(* IEC 61131-3 sources: llm-plc-st-eval/data/definitivo/gemini-3.1-pro-preview/I4/zero_shot, 3 files *)

(* ---- ejec_1.st ---- *)
```iecst
FUNCTION_BLOCK FB_EstrellaTriangulo
VAR_INPUT
    btnMarcha : BOOL; // Botón de arranque
    btnParo   : BOOL; // Botón de parada (prioridad a la parada)
END_VAR

VAR_OUTPUT
    kM : BOOL; // Contactor principal
    kY : BOOL; // Contactor de estrella
    kD : BOOL; // Contactor de triángulo
END_VAR

VAR
    tonEstrella   : TON; // Temporizador para la fase de estrella (8s)
    tonTransicion : TON; // Temporizador para el tiempo muerto (100ms)
END_VAR

// 1. Lógica del contactor principal (kM)
// Enclavamiento con btnMarcha, se rompe al pulsar btnParo
kM := (btnMarcha OR kM) AND NOT btnParo;

// 2. Temporizadores
// El temporizador de estrella inicia al arrancar el motor (kM = TRUE)
tonEstrella(IN := kM, PT := T#8S);

// El temporizador de transición inicia cuando termina la fase de estrella
tonTransicion(IN := tonEstrella.Q, PT := T#100MS);

// 3. Lógica de los contactores de fase (con enclavamiento mutuo de seguridad)
// kY se activa con kM, se apaga al terminar tonEstrella, y nunca si kD está activo
kY := kM AND NOT tonEstrella.Q AND NOT kD;

// kD se activa al terminar el tiempo muerto, y nunca si kY está activo
kD := kM AND tonTransicion.Q AND NOT kY;

END_FUNCTION_BLOCK
```

(* ---- ejec_2.st ---- *)
```iecst
FUNCTION_BLOCK FB_EstrellaTriangulo
VAR_INPUT
    btnMarcha : BOOL; (* Botón de inicio del motor *)
    btnParo   : BOOL; (* Botón de parada del motor *)
END_VAR

VAR_OUTPUT
    kM : BOOL; (* Contactor principal *)
    kY : BOOL; (* Contactor de estrella *)
    kD : BOOL; (* Contactor de triángulo *)
END_VAR

VAR
    xEnMarcha   : BOOL; (* Memoria de estado del motor *)
    tonEstrella : TON;  (* Temporizador para la fase de estrella *)
    tonTrans    : TON;  (* Temporizador para el tiempo muerto (transición) *)
END_VAR

(* Lógica de retención (Marcha / Paro) *)
IF btnParo THEN
    xEnMarcha := FALSE;
ELSIF btnMarcha THEN
    xEnMarcha := TRUE;
END_IF;

(* Temporizador de la fase Estrella (8 segundos) *)
tonEstrella(IN := xEnMarcha, PT := T#8S);

(* Temporizador de tiempo muerto entre Estrella y Triángulo (100 ms) *)
(* Inicia cuando termina la fase de estrella *)
tonTrans(IN := tonEstrella.Q, PT := T#100MS);

(* Asignación de salidas con enclavamientos de seguridad *)
(* El contactor principal se activa siempre que el sistema esté en marcha *)
kM := xEnMarcha;

(* Estrella: Activo en marcha, antes de los 8s, y NUNCA si Triángulo está activo *)
kY := xEnMarcha AND NOT tonEstrella.Q AND NOT kD;

(* Triángulo: Activo en marcha, tras el tiempo muerto, y NUNCA si Estrella está activo *)
kD := xEnMarcha AND tonTrans.Q AND NOT kY;

END_FUNCTION_BLOCK
```

(* ---- ejec_3.st ---- *)
```iecst
FUNCTION_BLOCK FB_EstrellaTriangulo
VAR_INPUT
    btnMarcha : BOOL; // Botón de arranque
    btnParo   : BOOL; // Botón de parada (TRUE = detener)
END_VAR

VAR_OUTPUT
    kM : BOOL; // Contactor principal
    kY : BOOL; // Contactor de estrella
    kD : BOOL; // Contactor de triángulo
END_VAR

VAR
    bRun        : BOOL; // Memoria del estado de marcha
    tonStar     : TON;  // Temporizador para la fase de estrella
    tonDeadTime : TON;  // Temporizador para el tiempo muerto
END_VAR

// 1. Lógica de retención (Marcha / Paro)
// El paro tiene prioridad sobre la marcha
IF btnParo THEN
    bRun := FALSE;
ELSIF btnMarcha THEN
    bRun := TRUE;
END_IF;

// 2. Temporizador de la fase de estrella (8 segundos)
tonStar(IN := bRun, PT := T#8S);

// 3. Control del contactor de Estrella (kY)
// Activo si hay marcha, no ha terminado el tiempo de estrella y kD está apagado (enclavamiento)
kY := bRun AND NOT tonStar.Q AND NOT kD;

// 4. Temporizador de tiempo muerto (100 milisegundos)
// Comienza a contar solo cuando termina la fase de estrella y kY se ha desactivado
tonDeadTime(IN := tonStar.Q AND NOT kY, PT := T#100MS);

// 5. Control del contactor de Triángulo (kD)
// Activo si hay marcha, terminó el tiempo muerto y kY está apagado (enclavamiento)
kD := bRun AND tonDeadTime.Q AND NOT kY;

// 6. Control del contactor Principal (kM)
// Activo siempre que el sistema esté en marcha
kM := bRun;

END_FUNCTION_BLOCK
```
